(* IEC 61131-3 sources: rusty/compiler/plc_cfc/fixtures/blocks/valid/program_chain, 1 file *)

(* ---- callees.st ---- *)
PROGRAM counter
VAR_INPUT
    in : DINT;
END_VAR
VAR_OUTPUT
    out : DINT;
END_VAR
    out := out + in;
END_PROGRAM

PROGRAM doubler
VAR_INPUT
    in : DINT;
END_VAR
VAR_OUTPUT
    out : DINT;
END_VAR
    out := in * 2;
END_PROGRAM
